{attribute 'qualified_only'}
VAR_GLOBAL
	aKistlerOut AT %Q* : ARRAY[0..199] OF BYTE; // PLC -> maXYmos
    aKistlerIn  AT %I* : ARRAY[0..199] OF BYTE; // maXYmos -> PLC
	
	bKistlerSafetyEnableOK AT %I* : BOOL; //kistler safety
	
	
END_VAR

(* stored: Version 1.1.0.1
   GVL GVL_KISTLER_IO: Id {613015f5-64b5-41ad-bf74-99e71be07f06} *)
